// LS Electric XG5000 project: NewPLC
// PLC LSPLC
// module base 0 slot 0: 입력 모듈:XGI-D24A/B (DC 24V 입력, 32점 (전류소스 싱크공용/ 전류소스 입력))
// module base 0 slot 1: 출력 모듈:XGQ-TR4A/B (트랜지스터 출력, 32점 (0.1A용, 싱크출력/소스출력))
// module base 0 slot 2: 위치결정 모듈:XGF-PN4B (위치결정 EtherCAT 네트워크 표준형, 4축)

PROGRAM NewProgram (task: 스캔 프로그램)

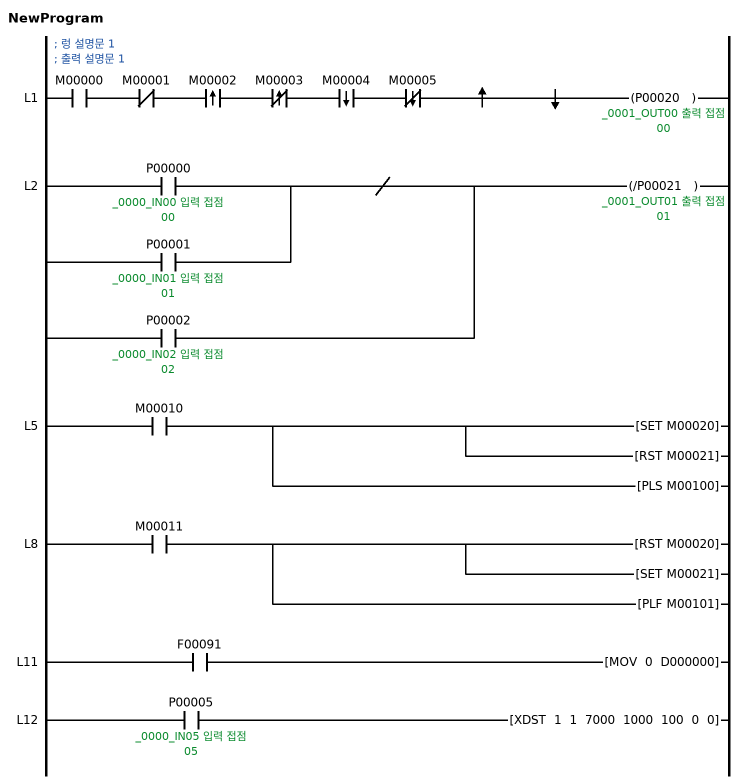
// 렁 설명문 1
; L1
LOAD      M00000
AND NOT   M00001
ANDP      M00002
ANDP NOT  M00003
ANDN      M00004
ANDN NOT  M00005
R_EDGE
F_EDGE
OUT       P00020	// _0001_OUT00 출력 접점 00
// output comment: 출력 설명문 1
; L2
LOAD      P00000	// _0000_IN00 입력 접점 00
OR        P00001	// _0000_IN01 입력 접점 01
NOT
OR        P00002	// _0000_IN02 입력 접점 02
OUT NOT   P00021	// _0001_OUT01 출력 접점 01
; L5
LOAD      M00010
SET       M00020
RST       M00021
OUTP      M00100
; L8
LOAD      M00011
RST       M00020
SET       M00021
OUTN      M00101
; L11
LOAD      F00091
MOV       0 D000000
; L12
LOAD      P00005	// _0000_IN05 입력 접점 05
XDST      1 1 7000 1000 100 0 0